// TIA Portal V21 export
// export: Created 2000-01-01T00:00:00.0000000Z, ExportSetting None
TYPE "UDT_HMI_CylinderCtrl"
   STRUCT
      bManualMode { ExternalWritable := 'False'} : Bool;   // TRUE: 手动模式, FALSE: 自动模式
      bManualExtendCmd { ExternalWritable := 'False'} : Bool;   // HMI手动伸出触发
      bManualRetractCmd { ExternalWritable := 'False'} : Bool;   // HMI手动缩回触发
      bResetCmd { ExternalWritable := 'False'} : Bool;   // HMI故障复位按钮
      tTimeoutSV { ExternalWritable := 'False'} : Time;   // 动作超时设定值（默认 T#3s）
      bIsExtended { ExternalWritable := 'False'} : Bool;   // 状态反馈：伸出到位
      bIsRetracted { ExternalWritable := 'False'} : Bool;   // 状态反馈：缩回到位
      bValveExtendOut { ExternalWritable := 'False'} : Bool;   // 状态反馈：伸出阀输出状态
      bValveRetractOut { ExternalWritable := 'False'} : Bool;   // 状态反馈：缩回阀输出状态
      bFault { ExternalWritable := 'False'} : Bool;   // 状态反馈：综合故障标志
      wStatus { ExternalWritable := 'False'} : Word;   // 状态码：16#0000正常, 16#8401伸出超时, 16#8402缩回超时, 16#8403前后磁性开关同时亮, 16#8404急停切断
   END_STRUCT;
END_TYPE
